Fanuc KAREL source: kt00371.KL

-- PROVISIONAL review KL for V770-1; original PC SHA256 535ea3db986bdea48e0c6c8cadcc1aeb1b5f29d7e525e72a0141922ae1b5df44
-- Incomplete behavior may be omitted. Consult companion uncertainty JSON. Do not deploy.
PROGRAM KT00371
%NOLOCKGROUP
VAR
  R1 : REAL
  OUT : BOOLEAN
-- UNRESOLVED_DECL Y2 type=002018
BEGIN
  -- UNRESOLVED_PC offsets 5-16; opcodes 2E,23
  -- UNRESOLVED_PC offsets 21-35; opcodes 2E,22,9D,33,B2
  -- UNRESOLVED_PC offsets 40-63; opcodes 21,22,9D,33,B1,64,70,23
  -- UNRESOLVED_PC offsets 68-72; opcodes 7F
END KT00371
